GLOBALCONSTANTS OpcString (* OPC-UA-IDs fuer STRING ueber CAN (Uebungen 137c, 139c) *)
  (* Standard: 61499-1; Description: Copyright (c) 2026 Meisterschulen am Ostbahnhof This program and the accompanying materials are made available under the terms of the Eclipse Public License 2.0 which is available at https://www.eclipse.org/legal/epl-2.0/ SPDX-License-Identifier: EPL-2.0 *)
  (* Version 1.0, 2026-11-14, Franz Höpfinger, Meisterschulen am Ostbahnhof, Empfangener Text lokal per PUBLISH (WRITE) *)
  PACKAGE Uebungen::const::Uebung_130_139;
  VAR_GLOBAL CONSTANT
    U137_TEXT_NODE : WSTRING := "/Objects/Uebungen/U137/Text,1:s=U137_Text"; (* 137c: Knoten Text *)
    U137_TEXT_WRITE : WSTRING := MyLib_OPC::F_OPC_LOCAL("WRITE", U137_TEXT_NODE); (* 137c: Text lokal schreiben *)
    U139_TEXT_NODE : WSTRING := "/Objects/Uebungen/U139/Text,1:s=U139_Text"; (* 139c: Knoten Text *)
    U139_TEXT_WRITE : WSTRING := MyLib_OPC::F_OPC_LOCAL("WRITE", U139_TEXT_NODE); (* 139c: Text lokal schreiben *)
  END_VAR
END_GLOBALCONSTANTS
